(* IEC 61131-3 sources: llm-plc-st-eval/data/definitivo/gpt-4o-2024-08-06/I6/zero_shot, 3 files *)

(* ---- ejec_1.st ---- *)
```pascal
FUNCTION_BLOCK FB_Temperatura
VAR_INPUT
    rawTemp : INT; // Valor de entrada de temperatura en bruto
END_VAR

VAR_OUTPUT
    tempC : REAL; // Temperatura calculada en grados Celsius
    enfriador : BOOL; // Estado del enfriador
    almSensor : BOOL; // Alarma de sensor
END_VAR

VAR
    tempC_prev : REAL; // Almacena el valor anterior de tempC para histéresis
END_VAR

// Constantes para la conversión de la señal de entrada a grados Celsius
CONST
    SCALE_FACTOR : REAL := 100.0 / 27648.0; // Factor de escala para convertir rawTemp a grados Celsius
END_CONST

// Cuerpo del bloque de función
BEGIN
    // Verificar si rawTemp está fuera de rango
    IF (rawTemp < 0) OR (rawTemp > 27648) THEN
        almSensor := TRUE; // Activar alarma de sensor
        enfriador := FALSE; // Desactivar enfriador
    ELSE
        almSensor := FALSE; // Desactivar alarma de sensor
        // Convertir rawTemp a grados Celsius
        tempC := rawTemp * SCALE_FACTOR;

        // Control del enfriador con histéresis
        IF tempC >= 80.0 THEN
            enfriador := TRUE; // Activar enfriador
        ELSIF tempC <= 75.0 THEN
            enfriador := FALSE; // Desactivar enfriador
        ELSE
            // Mantener el estado anterior del enfriador
            enfriador := enfriador;
        END_IF;
    END_IF;
END_FUNCTION_BLOCK
```

(* ---- ejec_2.st ---- *)
```pascal
FUNCTION_BLOCK FB_Temperatura
VAR_INPUT
    rawTemp : INT; // Entrada de la señal de temperatura cruda
END_VAR

VAR_OUTPUT
    tempC : REAL; // Salida de la temperatura en grados Celsius
    enfriador : BOOL; // Estado del enfriador
    almSensor : BOOL; // Alarma de sensor
END_VAR

VAR
    tempC_prev : REAL; // Variable para almacenar el valor anterior de tempC
END_VAR

// Conversión de la señal cruda a grados Celsius
tempC := (REAL(rawTemp) / 27648.0) * 100.0;

// Comprobación de límites de la señal cruda
IF (rawTemp < 0) OR (rawTemp > 27648) THEN
    almSensor := TRUE; // Activar alarma de sensor
    enfriador := FALSE; // Desactivar enfriador
ELSE
    almSensor := FALSE; // Desactivar alarma de sensor

    // Control del enfriador con histéresis
    IF tempC >= 80.0 THEN
        enfriador := TRUE; // Activar enfriador
    ELSIF tempC <= 75.0 THEN
        enfriador := FALSE; // Desactivar enfriador
    ELSE
        // Mantener el estado actual del enfriador
        enfriador := enfriador;
    END_IF
END_IF
END_FUNCTION_BLOCK
```

(* ---- ejec_3.st ---- *)
```pascal
FUNCTION_BLOCK FB_Temperatura
VAR_INPUT
    rawTemp : INT; // Valor de entrada de temperatura cruda
END_VAR

VAR_OUTPUT
    tempC : REAL; // Temperatura calculada en grados Celsius
    enfriador : BOOL; // Estado del enfriador
    almSensor : BOOL; // Alarma de sensor
END_VAR

VAR
    tempC_prev : REAL; // Valor previo de tempC para histéresis
END_VAR

// Conversión de rawTemp a grados Celsius
tempC := (REAL(rawTemp) * 100.0) / 27648.0;

// Comprobación de límites de rawTemp
IF (rawTemp < 0) OR (rawTemp > 27648) THEN
    almSensor := TRUE; // Activar alarma de sensor
    enfriador := FALSE; // Desactivar enfriador
ELSE
    almSensor := FALSE; // Desactivar alarma de sensor

    // Control del enfriador con histéresis
    IF tempC >= 80.0 THEN
        enfriador := TRUE; // Activar enfriador
    ELSIF tempC <= 75.0 THEN
        enfriador := FALSE; // Desactivar enfriador
    ELSE
        // Mantener el estado anterior del enfriador
        enfriador := enfriador;
    END_IF
END_IF
END_FUNCTION_BLOCK
```
